(* IEC 61131-3 sources: nautilus/website/lessons/b4-counter/variants/bad-full-at-four, 1 file *)

(* ---- program.st ---- *)
PROGRAM Counter
VAR
    parcels : CTU;   (* counts, and says when it has reached its preset *)
END_VAR

parcels(CU := Eye, R := Reset, PV := 4);   (* counts each rising edge of Eye *)

Count := parcels.CV;
Full  := parcels.Q;
END_PROGRAM
